(* IEC 61131-3 sources: Lasal-MCP/examples/SampleSource/LASALScreenAdvancedSolution/LASALScreenAdvancedSolution/LASALScreenAdvacnedSolution/Stations/Terminal/HMI/Class/MyColorBar, 1 file *)

(* ---- MyColorBar.st ---- *)
(*!
<Class
	Name               = "MyColorBar"
	Revision           = "0.0"
	RealtimeTask       = "false"
	CyclicTask         = "false"
	BackgroundTask     = "false"
	Sigmatek           = "false"
	OSInterface        = "false"
	HighPriority       = "false"
	Automatic          = "false"
	UpdateMode         = "Prescan"
	SharedCommandTable = "true"
	Objectsize         = "(480,240)">
	<Channels>
		<Server Name="IntError" Visualized="false" Initialize="false" WriteProtected="true" Retentive="false"/>
		<Client Name="_Grafix" Required="false" Internal="false"/>
		<Client Name="SigCLib" Required="false" Internal="false"/>
	</Channels>
	<Network Name="MyColorBar">
		<!-- List of Components in this network -->
		<Components>
			<Object
				Name       = "_base"
				Class      = "_MyIO"
				Position   = "(218,120)"
				Visualized = "true"
				Remotely   = "true">
				<Channels>
					<Server Name="Refresh"/>
					<Server Name="Server0"/>
					<Client Name="Graphic"/>
					<Client Name="Lse"/>
				</Channels>
			</Object>
		</Components>
		<Comments>
		</Comments>
		<!-- List of Connections in this network -->
		<Connections>
			<Connection Source="this.Server0" Destination="_base.Server0" Vertices="(706,210),(534,210),"/>
			<Connection Source="this.Refresh" Destination="_base.Refresh" Vertices="(706,270),(534,270),"/>
			<Connection Source="_base.Lse" Destination="this.Lse" Vertices="(218,210),(38,210),"/>
		</Connections>
		<!-- Headerfiles -->
		<Options>
		</Options>
	</Network>
</Class>
*)
#pragma using _MyIO

MyColorBar : CLASS
: _MyIO
  //Servers:
	IntError 	: SvrCh_DINT;
  //Clients:
	_Grafix 	: CltChCmd__Grafix;
	SigCLib 	: CltChCmd_SigCLib;
  //Variables:
		BarHeight 	: DINT;
		MinLimit 	: DINT;
		MaxLimit 	: DINT;
		MinBorder 	: DINT;
		MaxBorder 	: DINT;
		ActValue 	: DINT;
		ShowValue 	: BOOL;
		MinColor 	: UDINT;
		BarColor 	: UDINT;
		MaxColor 	: UDINT;
		pUnit 	: ^_CHAR;
		ActPixel 	: DINT;
		LowerSpaceHeight 	: INT;
		UpperSpaceHeight 	: INT;
		LowerSpace 	: _ROOM;
		MidSpace 	: _ROOM;
		UpperSpace 	: _ROOM;
		pError 	: ^CHAR;
  //Functions:
				//! <Function Comment="this method is called everytime when system wants to redraw the io" Name="Draw"/>
	FUNCTION __CDECL VIRTUAL GLOBAL Draw
		VAR_INPUT
			pio 	: ^_IO;			//! <Variable Comment="pointer to _IO information" Name="Draw.pio"/>
			pr 	: ^_RESULT;			//! <Variable Comment="pointer to _RESULT information" Name="Draw.pr"/>
			pv 	: ^_VARIABLE;			//! <Variable Comment="pointer to io _VARIABLE information" Name="Draw.pv"/>
			input 	: BOOL;			//! <Variable Comment="TRUE it&apos;s an input&#13;&#10;FALSE it&apos;s an output" Name="Draw.input"/>
		END_VAR
		VAR_OUTPUT
			retcode (EAX) 	: _DOIT;			//! <Variable Comment="for the returnstatement there are 3 different possibilities&#13;&#10;  _IDLE ..... the system should goon like it is (system goes on)&#13;&#10;  _IDIDIT ... i did it (system is ready)&#13;&#10;  _IFAILED .. i tried to do my best, but i failed (system is re" Name="Draw.retcode"/>
		END_VAR;
				//! <Function Comment="this method is called everytime when system wants to get data for defined io.&#13;&#10;&#13;&#10;pr ........ &#13;&#10;pio ....... pointer to io information&#13;&#10;pv ........ pointer to io variableinformation&#13;&#10;input ..... TRUE it&apos;s an input / FALSE it&apos;s an output&#13;&#10;&#13;&#10;for the returnstatement there are 3 different possibilities&#13;&#10;_IDLE ..... the system should goon like it is (system goes on)&#13;&#10;_IDIDIT ... i did it (system is ready)&#13;&#10;_IFAILED .. i tried to do my best, but i failed (system is ready)&#13;&#10;&#13;&#10;if you want to do it let&apos;s return _IDIDIT and initialize the  structure _RESULT&#13;&#10;" Name="GetData"/>
	FUNCTION __CDECL VIRTUAL GLOBAL GetData
		VAR_INPUT
			pr 	: ^_RESULT;			//! <Variable Comment="pointer to _RESULT information" Name="GetData.pr"/>
			pio 	: ^_IO;			//! <Variable Comment="pointer to _IO information" Name="GetData.pio"/>
			pv 	: ^_VARIABLE;			//! <Variable Comment="pointer to _VARIABLE information given by LSE" Name="GetData.pv"/>
			input 	: BOOL;			//! <Variable Comment="TRUE it&apos;s an input&#13;&#10;FALSE it&apos;s an output" Name="GetData.input"/>
		END_VAR
		VAR_OUTPUT
			retcode (EAX) 	: _DOIT;			//! <Variable Comment="for the returnstatement there are 3 different possibilities&#13;&#10;  _IDLE ..... the system should goon like it is (system goes on)&#13;&#10;  _IDIDIT ... i did it (system is ready)&#13;&#10;  _IFAILED .. i tried to do my best, but i failed (system is ready)" Name="GetData.retcode"/>
		END_VAR;
				//! <Function Comment="this method is called once right in front of drawing the object.&#13;&#10;for example open screen&#13;&#10;" Name="IF_Start"/>
	FUNCTION __CDECL VIRTUAL GLOBAL IF_Start
		VAR_INPUT
			pio 	: ^_IO;			//! <Variable Comment="pointer to _IO information" Name="IF_Start.pio"/>
			firsttime 	: BOOL;			//! <Variable Comment="true: when system wants to view drawing after open screen&#13;&#10;false: when system wants to redraw background" Name="IF_Start.firsttime"/>
		END_VAR;
  //Tables:
	FUNCTION @STD
		VAR_OUTPUT
			ret_code	: CONFSTATES;
		END_VAR;
	FUNCTION GLOBAL TAB @CT_;
END_CLASS;

#pragma usingLtd _Grafix
#pragma usingLtd SigCLib

FUNCTION __CDECL VIRTUAL GLOBAL MyColorBar::IF_Start
	VAR_INPUT
		pio 	: ^_IO;
		firsttime 	: BOOL;
	END_VAR

  if (firsttime = TRUE) then
    BarHeight := (pio^.space.xy2.y - pio^.space.xy1.y) + 1;
  end_if;

END_FUNCTION

FUNCTION __CDECL VIRTUAL GLOBAL MyColorBar::GetData
	VAR_INPUT
		pr 	: ^_RESULT;
		pio 	: ^_IO;
		pv 	: ^_VARIABLE;
		input 	: BOOL;
	END_VAR
	VAR_OUTPUT
		retcode (EAX) 	: _DOIT;
	END_VAR
  VAR
  	varno : UDINT;
    plabel : ^_VARLABEL;
  END_VAR

  retcode := _IFAILED;

  // check for valid pointer to udc
  if (pio^.theurge <> NIL) then

    // check no of data parameters
    if (pio^.theurge^.memvarlabel.no = 6) then

      // get pointer to first datasource of the udc
      plabel := pio^.theurge^.memvarlabel.ptr;

      // write value to variable
      VarList_GetValue(p0:= plabel,
                       p1:= #MinLimit,
                       x2:= FALSE);

      // increase pointer to label and write next variable
      plabel += sizeof(_VARLABEL);
      VarList_GetValue(p0:= plabel,
                       p1:= #MaxLimit,
                       x2:= FALSE);

      // increase pointer to label and write next variable
      plabel += sizeof(_VARLABEL);
      VarList_GetValue(p0:= plabel,
                       p1:= #MinBorder,
                       x2:= FALSE);

      // increase pointer to label and write next variable
      plabel += sizeof(_VARLABEL);
      VarList_GetValue(p0:= plabel,
                       p1:= #MaxBorder,
                       x2:= FALSE);

      // increase pointer to label and write next variable
      plabel += sizeof(_VARLABEL);
      VarList_GetValue(p0:= plabel,
                       p1:= #ActValue,
                       x2:= FALSE);

      // get no of selected Server
      varno := to_udint(plabel^.info[0].value);

      // get pointer to unit text
      pUnit := VarList_GetTextByNo(x0:= varno,
                                   x1:= 5);

      // increase pointer to label and write next variable
      plabel += sizeof(_VARLABEL);
      VarList_GetValue(p0:= plabel,
                       p1:= #ShowValue$DINT,
                       x2:= FALSE);

      // get colors
      MinColor := pio^.theurge^.memcolor.ptr^;
      BarColor := (pio^.theurge^.memcolor.ptr + sizeof(_COLOR))^;
      MaxColor := (pio^.theurge^.memcolor.ptr + (2 * sizeof(_COLOR)))^;

      // switch of cablebreak
      if (ActValue < 0) then
        ActValue := MaxLimit;
      end_if;

      // calculate actual Pixel height
      ActPixel := to_dint((to_real(BarHeight) / to_real(MaxLimit)) * to_real(ActValue));

      // calculate height lower- and UpperSpace
      LowerSpaceHeight := to_int(DIV_AB_BY_C(A:= BarHeight,
                                             B:= MinBorder,
                                             _C:= MaxLimit));

      UpperSpaceHeight := to_int(DIV_AB_BY_C(A:= BarHeight,
                                             B:= MaxBorder,
                                             _C:= MaxLimit));
      // set koords from spaces
      LowerSpace.xy1.x := pio^.space.xy1.x;
      LowerSpace.xy1.y := pio^.space.xy2.y - LowerSpaceHeight;
      LowerSpace.xy2.x := pio^.space.xy2.x;
      LowerSpace.xy2.y := pio^.space.xy2.y;

      MidSpace.xy1.x := pio^.space.xy1.x;
      MidSpace.xy1.y := pio^.space.xy2.y - UpperSpaceHeight;
      MidSpace.xy2.x := pio^.space.xy2.x;
      MidSpace.xy2.y := pio^.space.xy2.y - LowerSpaceHeight;

      UpperSpace.xy1.x := pio^.space.xy1.x;
      UpperSpace.xy1.y := pio^.space.xy1.y;
      UpperSpace.xy2.x := pio^.space.xy2.x;
      UpperSpace.xy2.y := pio^.space.xy2.y - UpperSpaceHeight;

      // set pixel height
      pr^.value := ActPixel;

      retcode := _IDIDIT;

    else
      IntError := -2; // invalid data parameter no
      return;

    end_if;
  else
    IntError := -1; // invalid pointer
    return;
  end_if;

END_FUNCTION

FUNCTION __CDECL VIRTUAL GLOBAL MyColorBar::Draw
	VAR_INPUT
		pio 	: ^_IO;
		pr 	: ^_RESULT;
		pv 	: ^_VARIABLE;
		input 	: BOOL;
	END_VAR
	VAR_OUTPUT
		retcode (EAX) 	: _DOIT;
	END_VAR
  VAR
    act : _NEWSCREEN;
    text : array[0..19] of char;
  END_VAR

  // switch to offscreen
  push_screen(p0:=#act);

  // Copy content of the current screen to the offscreen.
  _Grafix.PutImage(image:=#pio^.image, x0:=DEFKOORD, y0:=DEFKOORD);

  // draw background
  _Grafix.Beam(x0:= pio^.space.xy1.x,
               y0:= pio^.space.xy1.y,
               x1:= pio^.space.xy2.x,
               y1:= pio^.space.xy2.y,
               attrib:= pio^.attrib,
               color:= pio^.colback);

  // draw lower space with actual value
  if (ActPixel <= LowerSpaceHeight) then

    color_course(p0:= #LowerSpace,
                 x1:= to_int(ActPixel) * -1,
                 x2:= MinColor,
                 x3:= BarColor,
                 x4:= T_COPY or T_SOLID or T_VERTBOUND);

  // draw lower space with max height
  else
    color_course(p0:= #LowerSpace,
                 x1:= LowerSpaceHeight * -1,
                 x2:= MinColor,
                 x3:= BarColor,
                 x4:= T_COPY or T_SOLID or T_VERTBOUND);
  end_if;

  // draw midSpace with actual value
  if ((ActPixel > LowerSpaceHeight) & (ActPixel < UpperSpaceHeight)) then

    _Grafix.Beam(x0:= MidSpace.xy1.x,
                 y0:= MidSpace.xy2.y - (to_int(ActPixel) - LowerSpaceHeight),
                 x1:= MidSpace.xy2.x,
                 y1:= MidSpace.xy2.y,
                 attrib:= T_COPY or T_SOLID or T_VERTBOUND,
                 color:= BarColor);

  // draw upperspace and MidSpace with max height
  elsif (ActPixel >= UpperSpaceHeight) then

    _Grafix.Beam(x0:= MidSpace.xy1.x,
                 y0:= MidSpace.xy1.y,
                 x1:= MidSpace.xy2.x,
                 y1:= MidSpace.xy2.y,
                 attrib:= T_COPY or T_SOLID or T_VERTBOUND,
                 color:= BarColor);

    color_course(p0:= #UpperSpace,
                 x1:= (to_int(ActPixel) - UpperSpaceHeight) * -1,
                 x2:= BarColor,
                 x3:= MaxColor,
                 x4:= T_COPY or T_SOLID or T_VERTBOUND);
  end_if;

  if (ShowValue = TRUE) then

    DToA(p0:= #text[0],
         x1:= ActValue,
         x2:= 16#0800,
         x3:= sizeof(_ASCII));

    pError := SigCLib.StrCat(ps1:= #text[0],
                             ps2:= " ");

    if (pError <> #text[0]) then
      IntError := -3;
      return;
    end_if;

    // StrCat to copy the Unicode Unit from LSE
    StrCat(p0:= #text[0],
           x1:= sizeof(_ASCII),
           p2:= pUnit,
           x3:= sizeof(_UNI));

    OutTextAlign(p0:= #text[0],
                 x1:= 0,
                 p1:= #pio^.space,
                 x2:= pio^.font,
                 x3:= pio^.attrib,
                 x9:= pio^.frametype,
                 x4:= pio^.coltxt,
                 x5:= _Grafix.MakeColor(backcolor:=INVISIBLE, frontcolor:=INVISIBLE),
                 x6:= _Grafix.MakeColor(backcolor:=INVISIBLE, frontcolor:=INVISIBLE),
                 x7:= sizeof(_ASCII));
  end_if;

  // visible screen switched on
  pop_screen(p0:= #act);

  // copy image on visible screen
  copy_screen(p0:= #act, p1:= #pio^.space);

  retcode := _IDIDIT;

END_FUNCTION
